{attribute 'qualified_only'}
{attribute 'strict'}
{attribute 'to_string'}
TYPE E_BB_States :
(
	Unknown	:= 0,
	OUT		:= 1,
	IN		:= 2
) UINT;
END_TYPE

(* stored: Version 1.1.0.1
   DUT E_BB_States: Id {3f522ed9-7d8a-45e5-97f2-fc34f5b8fa18} *)
